Fanuc KAREL source: kb00129.KL

PROGRAM KB00129
%STACKSIZE=65535
%PRIORITY=65535
%NOLOCKGROUP
VAR
P1 : STRING[80]
P2 : BOOLEAN
P3 : BOOLEAN
P4 : INTEGER
BEGIN
P1='A'
P2=TRUE
P3=TRUE
P4=1
PAUSE_TASK(P1,P2,P3,P4)
END KB00129
